// TIA Portal V18 export
VAR_GLOBAL   // PLC tag table "BYPASS_APERTADEIRAS"
   start AT %I1500.1 : Bool;
   remover AT %I1500.2 : Bool;
   reset AT %I1500.3 : Bool;
   MOD1_OK AT %Q1594.0 : Bool;
   MOD2_OK AT %Q1594.1 : Bool;
   RESET_MOD_1 AT %M9.1 : Bool;
   RESET_MOD_2 AT %M9.2 : Bool;
   VALIDACA0_MOD1 AT %M9.6 : Bool;
   VALIDAÇÃO_MOD2 AT %M12.0 : Bool;
   VALIDACAO_ANDON_MOD2 AT %M12.2 : Bool;
   VALIDACAO_ANDON_MOD1 AT %M12.3 : Bool;
   LEANDRO AT %M12.4 : Bool;
   BYPASS_ABST_OLEO AT %M12.6 : Bool;
   BYPASS_ABSTECIMENTO_OLEO AT %M12.7 : Bool;
   BYPASS_ESTANQ_CIL AT %M13.0 : Bool;
   BYPASS_SUP_FREIO AT %M2.1 : Bool;
   BYPASS_PY_EXCENTRICO AT %M2.2 : Bool;
   BYPASS_AP_HARPA AT %M12.5 : Bool;
   BYPASS_BUJAO AT %M13.1 : Bool;
   BYPASS_AP_BUJAO AT %M13.2 : Bool;
   BYPASS_TUBO_RPX AT %M13.3 : Bool;
   BYPASS_AP_TUBO_RPX AT %M13.4 : Bool;
   BYPASS_MOLA_HARPA AT %M13.5 : Bool;
   BYPASS_CARCACA AT %M13.6 : Bool;
   BYPASS_AP_CARCA AT %M13.7 : Bool;
   BYPASS_TALHA_DIF AT %M28.0 : Bool;
   BYPASS_SENSOR_TALHA_DIF AT %M28.1 : Bool;
   BYPASS_PYJUNTA AT %M28.2 : Bool;
   BYPASS_PY_JUNTA AT %M28.3 : Bool;
   BYPASS_CRAWFOOT AT %M28.4 : Bool;
   BYPASS_AP_CRAWFOOT AT %M28.5 : Bool;
   BYPASS_DUPLO_FUSO AT %M28.6 : Bool;
   BYPASS_AP_DUPLO_FUSO AT %M28.7 : Bool;
   BYPASS_P_ESCONDIDA AT %M29.0 : Bool;
   BYPASS_AP_PORCA_ESCON AT %M29.1 : Bool;
   BYPASS_SUP_CIL AT %M29.2 : Bool;
   BYPASS_AP_SUP_CIL AT %M29.3 : Bool;
   BYPASS_PORCA_CIL AT %M29.4 : Bool;
   BYPASS_AP_PORCA_CIL AT %M29.5 : Bool;
   BYPASS_AP_SUP_FREIO AT %M29.6 : Bool;
   BYPASS_PYEXCENTRICO AT %M29.7 : Bool;
   BYPASS_CUBO_DISC AT %M30.0 : Bool;
   BYPASS_PY_CUBO_DISC AT %M30.1 : Bool;
   BYPASS_HOLDER AT %M30.2 : Bool;
   BYPASS_AP_HOLDER AT %M30.3 : Bool;
   BYPASS_CALIPER AT %M30.4 : Bool;
   BYPASS_AP_CALPER AT %M30.5 : Bool;
   BYPASS_PYCUBO_TAMBOR AT %M30.6 : Bool;
   BYPASS_PY_CUBO_TAMBOR AT %M30.7 : Bool;
   BYPASS_HASTE_ALV AT %M31.0 : Bool;
   BYPASS_AP_HASTE_ALV AT %M31.1 : Bool;
   BYPASS_APCUBO AT %M31.2 : Bool;
   BYPASS_AP_CUBO AT %M31.3 : Bool;
   BYPASS_CRAVADOR AT %M31.4 : Bool;
   BYPASS_AP_CRAVADOR AT %M31.5 : Bool;
   BYPASS_INDICADOR AT %M31.6 : Bool;
   BYPASS_AP_INDICADOR AT %M31.7 : Bool;
   BYPASS_VALVULA AT %M32.0 : Bool;
   BYPASS_AP_VALVULA AT %M32.1 : Bool;
   BYPASS_HELGE AT %M32.2 : Bool;
   BYPASS_PY_HELGE AT %M32.3 : Bool;
   BYPASS_PORCA_TERMINAL AT %M32.4 : Bool;
   BYPASS_AP_PORCA_TERMINAL AT %M32.5 : Bool;
   BYPASS_FILTRO_OLEO AT %M32.6 : Bool;
   BYPASS_AP_FILTRO_OLEO AT %M32.7 : Bool;
   BYPASS_REDUCAO AT %M33.0 : Bool;
   BYPASS_AP_REDUCAO AT %M33.1 : Bool;
   BYPASS_FLANGE AT %M33.2 : Bool;
   BYPASS_AP_FLANGE AT %M33.3 : Bool;
   BYPASS_ESTANQ_CILINDRO AT %M33.4 : Bool;
   BYPASS_ESTANQ_CARC AT %M33.5 : Bool;
   BYPASS_ESTANQ_CARCACA AT %M33.6 : Bool;
   EMERG_CABINE_ACIONADA AT %M35.1 : Bool;
   BYPASS_VALVULA_P50 AT %M35.6 : Bool;
   BYPASS_TAMPA_CALIPER_1 AT %M36.0 : Bool;
   BYPASS_AP_VALVULA_P50 AT %M36.1 : Bool;
   TESTE_LEITOR AT %M42.4 : Bool;
   IG_CONTROL_T AT %M43.7 : Bool;
   ABORTA_P05 AT %M2.5 : Bool;
   ABORTA_JOB_P05 AT %M2.6 : Bool;
   TORQUE_ATLAS6000_P15 AT %MD48 : Real;
   PULSO_BORDA_BYPASS AT %M3.1 : Bool;
   BORDA_BYPASS_AP AT %M3.2 : Bool;
   TORQUE_DUPLO_FUSO1 AT %MD52 : Real;
   AUX_APDP AT %M3.4 : Bool;
   SIGNAL_LOST_POKA_JUNTA AT %M3.5 : Bool;
   aux_inicio_receita_pky_p30 AT %M3.7 : Bool;
   JOBOK_POKA_JUNTA_P30 AT %M4.0 : Bool;
   BYPASS_TORQUIMETRO_DIGITAL_1 AT %M4.1 : Bool;
   BYPASS_REULAGEM_ALAVANCA_1 AT %M4.5 : Bool;
   antecipa_expedicao AT %M4.6 : Bool;
   SIGINAL_LOST_PCUBO AT %M5.0 : Bool;
   pulso_teste AT %M5.7 : Bool;
   JOBDONE_ABSTECIMENTO_OLEO AT %M7.3 : Bool;
   SIGNAL_LOST_ABAST_OLEO AT %M7.4 : Bool;
   Bypass_oring_P100 AT %M7.5 : Bool;
   BYPASS_ORING_MAP_P100 AT %M8.1 : Bool;
   SIGNAL_LOST_ORING_MAP AT %M8.3 : Bool;
   InputAuxEdi AT %M8.7 : Bool;
   InputAuxEtr AT %M9.0 : Bool;
   SEM_JOB_PY_OLEO AT %M56.6 : Bool;
   JOB_PY_OLEO AT %M56.7 : Bool;
   JOBDONE_PY_GRAXA AT %M57.2 : Bool;
   Bypass_jidoka_filtro AT %M57.3 : Bool;
   BYPASS_JIDOKA_FILTRO_OLEO_P125 AT %M57.4 : Bool;
   Bypass_vaselina AT %M57.5 : Bool;
   JobOK_vaselina AT %M57.6 : Bool;
   BYpassVaselina AT %M57.7 : Bool;
   resetsinais AT %M58.0 : Bool;
   Bypass_apcilin_pneumatico AT %M58.2 : Bool;
   Bypass_apcilin_pneumaticoP105 AT %M58.3 : Bool;
END_VAR
